// Value of bMoveAbortPending after a reset (MONETcommon#56, #66 part 1). A reset drops the pending move commands; a move that
// is still running must not run on to its old target, so the abort stop of #84 goes on: one MC_Stop per moving axis (#96),
// no bStop (no operator stop), moving axes are not reset (0x4260, #84).
// TRUE only if an enabled axis is moving (also homing). Not during an error (the drives are off) and not while a park runs
// (its motion is wanted; bPark is kept by the reset). An axis stuck in Stopping without motion does not count: a reset must
// still get out of a hung abort stop.
FUNCTION F_ResetMoveAbort : BOOL
VAR_INPUT
	bError			: BOOL;
	bParkRunning	: BOOL;		// TCS_command = park
	bAzMoving		: BOOL;		// enabled AND (InMotion OR InRamp OR Homing), per axis
	bElMoving		: BOOL;
	bDrMoving		: BOOL;
END_VAR

F_ResetMoveAbort := NOT bError AND NOT bParkRunning AND (bAzMoving OR bElMoving OR bDrMoving);

END_FUNCTION

(* stored: Version 1.1.0.1, ProductVersion 3.1.4024.15
   POU F_ResetMoveAbort: Id {8b6f3a52-1c0e-4d7a-9a35-5e2d41c7f0b9}, SpecialFunc None *)
